                num nValue[3]
            mdesc mMdesc
            num nActionIndex = 42
            num nDelay
            num nMoveType = 1
            num nPercentage
            num nSigValue = 1
        pointRx pPointRx[2] = {x=93.576632, y=-409.183941, z=700.107773, rx=0.434495, ry=-1.660891, rz=-0.491266, shoulder=lefty, elbow=enegative, wrist=wpositive}
        string sID
      [45]
        bool bMarked
        jointRx jJointRx = {j1=-101.229016, j2=121.246473, j3=-113.173387, j4=191.93634, j5=7.483782, j6=-91.0959406}
        pointRx pInter
        paraItem pParaItem
          [0]
            bool bSafePoint
            ifItem iIfItem
              [0]
                bool bANDOR[2]
                num nSigIndex[3]
                num nSigType[3]
                num nValue[3]
            mdesc mMdesc
            num nActionIndex = 42
            num nDelay
            num nMoveType = 1
            num nPercentage
            num nSigValue = 1
        pointRx pPointRx[2] = {x=-57.556145, y=-477.506256, z=700.107677, rx=0.434341, ry=-1.659983, rz=-0.491216, shoulder=lefty, elbow=enegative, wrist=wpositive}
        string sID
      [46]
        bool bMarked
        jointRx jJointRx = {j1=-100.83359, j2=118.28296, j3=-99.234912, j4=184.924538, j5=18.376568, j6=-84.328027}
        pointRx pInter
        paraItem pParaItem
          [0]
            bool bSafePoint
            ifItem iIfItem
              [0]
                bool bANDOR[2]
                num nSigIndex[3]
                num nSigType[3]
                num nValue[3]
            mdesc mMdesc
            num nActionIndex = 42
            num nDelay
            num nMoveType = 1
            num nPercentage
            num nSigValue = 1
        pointRx pPointRx[2] = {x=-71.199798, y=-566.082474, z=700.128795, rx=0.430138, ry=-1.661253, rz=-0.490771, shoulder=lefty, elbow=enegative, wrist=wpositive}
        string sID
      [47]
        bool bMarked
        jointRx jJointRx = {j1=-96.744625, j2=116.717504, j3=-93.79165, j4=184.203052, j5=22.358435, j6=-87.631438}
        pointRx pInter
        paraItem pParaItem
          [0]
            bool bSafePoint
            ifItem iIfItem
              [0]
                bool bANDOR[2]
                num nSigIndex[3]
                num nSigType[3]
                num nValue[3]
            mdesc mMdesc
            num nActionIndex = 42
            num nDelay
            num nMoveType = 1
            num nPercentage
            num nSigValue = 1
        pointRx pPointRx[2] = {x=-34.726735, y=-600.68007, z=700.128795, rx=0.429673, ry=-1.659562, rz=-0.490424, shoulder=lefty, elbow=enegative, wrist=wpositive}
        string sID
      [48]
        bool bMarked
        jointRx jJointRx = {j1=-95.531794, j2=118.469763, j3=-99.931703, j4=185.21224, j5=18.0199205, j6=-89.914501}
        pointRx pInter
        paraItem pParaItem
          [0]
            bool bSafePoint
            ifItem iIfItem
              [0]
                bool bANDOR[2]
                num nSigIndex[3]
                num nSigType[3]
                num nValue[3]
            mdesc mMdesc
            num nActionIndex = 42
            num nDelay
            num nMoveType = 1
            num nPercentage
            num nSigValue = 1
        pointRx pPointRx[2] = {x=-18.573295, y=-564.69379, z=700.128759, rx=0.42985, ry=-1.65955, rz=-0.49045, shoulder=lefty, elbow=enegative, wrist=wpositive}
        string sID
      [49]
        bool bMarked
        jointRx jJointRx = {j1=-92.248565, j2=118.548585, j3=-100.229526, j4=185.345375, j5=17.897666, j6=-93.328956}
        pointRx pInter
        paraItem pParaItem
          [0]
            bool bSafePoint
            ifItem iIfItem
              [0]
                bool bANDOR[2]
                num nSigIndex[3]
                num nSigType[3]
                num nValue[3]
            mdesc mMdesc
            num nActionIndex = 42
            num nDelay
            num nMoveType = 1
            num nPercentage
            num nSigValue = 1
        pointRx pPointRx[2] = {x=13.638528, y=-562.185834, z=700.128755, rx=0.429526, ry=-1.658701, rz=-0.490292, shoulder=lefty, elbow=enegative, wrist=wpositive}
        string sID
      [50]
        bool bMarked
        jointRx jJointRx = {j1=-92.0110168, j2=115.175363, j3=-88.916981, j4=183.775747, j5=25.818301, j6=-91.878431}
        pointRx pInter
        paraItem pParaItem
          [0]
            bool bSafePoint
            ifItem iIfItem
              [0]
                bool bANDOR[2]
                num nSigIndex[3]
                num nSigType[3]
                num nValue[3]
            mdesc mMdesc
            num nActionIndex = 42
            num nDelay
            num nMoveType = 1
            num nPercentage
            num nSigValue = 1
        pointRx pPointRx[2] = {x=13.638517, y=-627.787273, z=700.128718, rx=0.430872, ry=-1.659586, rz=-0.490435, shoulder=lefty, elbow=enegative, wrist=wpositive}
        string sID
      [51]
        bool bMarked
        jointRx jJointRx = {j1=-97.374112, j2=108.454018, j3=-70.449442, j4=182.620747, j5=37.393534, j6=-85.196557}
        pointRx pInter
        paraItem pParaItem
          [0]
            bool bSafePoint
            ifItem iIfItem
              [0]
                bool bANDOR[2]
                num nSigIndex[3]
                num nSigType[3]
                num nValue[3]
            mdesc mMdesc
            num nActionIndex = 42
            num nDelay
            num nMoveType = 1
            num nPercentage
            num nSigValue = 1
        pointRx pPointRx[2] = {x=-56.645666, y=-719.0880848, z=700.128704, rx=0.430401, ry=-1.660167, rz=-0.490645, shoulder=lefty, elbow=enegative, wrist=wpositive}
        string sID
      [52]
        bool bMarked
        jointRx jJointRx = {j1=-97.840683, j2=111.886769, j3=-79.472132, j4=183.0096897, j5=31.798373, j6=-85.205581}
        pointRx pInter
        paraItem pParaItem
          [0]
            bool bSafePoint
            ifItem iIfItem
              [0]
                bool bANDOR[2]
                num nSigIndex[3]
                num nSigType[3]
                num nValue[3]
            mdesc mMdesc
            num nActionIndex = 42
            num nDelay
            num nMoveType = 1
            num nPercentage
            num nSigValue = 1
        pointRx pPointRx[2] = {x=-56.645667, y=-676.466244, z=700.128712, rx=0.429254, ry=-1.659449, rz=-0.490453, shoulder=lefty, elbow=enegative, wrist=wpositive}
        string sID
      [53]
        bool bMarked
        jointRx jJointRx = {j1=-99.139712, j2=112.699971, j3=-81.717312, j4=183.11065, j5=30.332067, j6=-84.0331021}
        pointRx pInter
        paraItem pParaItem
          [0]
            bool bSafePoint
            ifItem iIfItem
              [0]
                bool bANDOR[2]
                num nSigIndex[3]
                num nSigType[3]
                num nValue[3]
            mdesc mMdesc
            num nActionIndex = 42
            num nDelay
            num nMoveType = 1
            num nPercentage
            num nSigValue = 1
        pointRx pPointRx[2] = {x=-70.0879135, y=-664.155218, z=700.128714, rx=0.429183, ry=-1.659583, rz=-0.490504, shoulder=lefty, elbow=enegative, wrist=wpositive}
        string sID
      [54]
        bool bMarked
        jointRx jJointRx = {j1=-105.267989, j2=114.670594, j3=-87.395728, j4=183.340854, j5=26.462946, j6=-78.209203}
        pointRx pInter
        paraItem pParaItem
          [0]
            bool bSafePoint
            ifItem iIfItem
              [0]
                bool bANDOR[2]
                num nSigIndex[3]
                num nSigType[3]
                num nValue[3]
            mdesc mMdesc
            num nActionIndex = 42
            num nDelay
            num nMoveType = 1
            num nPercentage
            num nSigValue = 1
        pointRx pPointRx[2] = {x=-132.400518, y=-625.604431, z=700.128755, rx=0.42881, ry=-1.659576, rz=-0.490548, shoulder=lefty, elbow=enegative, wrist=wpositive}
        string sID
      [55]
        bool bMarked
        jointRx jJointRx = {j1=-104.169194, j2=109.68382, j3=-73.608878, j4=182.604541, j5=35.278725, j6=-78.44342}
        pointRx pInter
        paraItem pParaItem
          [0]
            bool bSafePoint
            ifItem iIfItem
              [0]
                bool bANDOR[2]
                num nSigIndex[3]
                num nSigType[3]
                num nValue[3]
            mdesc mMdesc
            num nActionIndex = 42
            num nDelay
            num nMoveType = 1
            num nPercentage
            num nSigValue = 1
        pointRx pPointRx[2] = {x=-137.458378, y=-695.112294, z=700.128753, rx=0.430847, ry=-1.65989, rz=-0.490478, shoulder=lefty, elbow=enegative, wrist=wpositive}
        string sID
      [56]
        bool bMarked
        jointRx jJointRx = {j1=-108.836483, j2=105.997726, j3=-64.330372, j4=182.193953, j5=40.744432, j6=-73.310916}
        pointRx pInter
        paraItem pParaItem
          [0]
            bool bSafePoint
            ifItem iIfItem
              [0]
                bool bANDOR[2]
                num nSigIndex[3]
                num nSigType[3]
                num nValue[3]
            mdesc mMdesc
            num nActionIndex = 42
            num nDelay
            num nMoveType = 1
            num nPercentage
            num nSigValue = 1
        pointRx pPointRx[2] = {x=-206.432129, y=-721.294628, z=700.128699, rx=0.4308, ry=-1.659754, rz=-0.490404, shoulder=lefty, elbow=enegative, wrist=wpositive}
        string sID
      [57]
        bool bMarked
        jointRx jJointRx = {j1=-117.384994, j2=111.318057, j3=-77.929976, j4=182.390665, j5=32.266362, j6=-65.120808}
        pointRx pInter
        paraItem pParaItem
          [0]
            bool bSafePoint
            ifItem iIfItem
              [0]
                bool bANDOR[2]
                num nSigIndex[3]
                num nSigType[3]
                num nValue[3]
            mdesc mMdesc
            num nActionIndex = 42
            num nDelay
            num nMoveType = 1
            num nPercentage
            num nSigValue = 1
        pointRx pPointRx[2] = {x=-282.767279, y=-630.359837, z=700.128774, rx=0.429, ry=-1.659295, rz=-0.490511, shoulder=lefty, elbow=enegative, wrist=wpositive}
        string sID
      [58]
        bool bMarked
        jointRx jJointRx = {j1=-126.0288968, j2=110.864642, j3=-76.715468, j4=182.00929387, j5=32.842378, j6=-56.143629}
        pointRx pInter
        paraItem pParaItem
          [0]
            bool bSafePoint
            ifItem iIfItem
              [0]
                bool bANDOR[2]
                num nSigIndex[3]
                num nSigType[3]
                num nValue[3]
            mdesc mMdesc
            num nActionIndex = 42
            num nDelay
            num nMoveType = 1
            num nPercentage
            num nSigValue = 1
        pointRx pPointRx[2] = {x=-377.367552, y=-587.693598, z=700.128774, rx=0.428889, ry=-1.659196, rz=-0.49055, shoulder=lefty, elbow=enegative, wrist=wpositive}
        string sID
      [59]
        bool bMarked
        jointRx jJointRx = {j1=-132.158352, j2=110.822497, j3=-76.606813, j4=181.740658, j5=32.799901, j6=-49.794511}
        pointRx pInter
        paraItem pParaItem
          [0]
            bool bSafePoint
            ifItem iIfItem
              [0]
                bool bANDOR[2]
                num nSigIndex[3]
                num nSigType[3]
                num nValue[3]
            mdesc mMdesc
            num nActionIndex = 42
            num nDelay
            num nMoveType = 1
            num nPercentage
            num nSigValue = 1
        pointRx pPointRx[2] = {x=-437.975867, y=-545.96373, z=700.144476, rx=0.425586, ry=-1.657208, rz=-0.495183, shoulder=lefty, elbow=enegative, wrist=wpositive}
        string sID
      [60]
        bool bMarked
        jointRx jJointRx = {j1=-130.472656, j2=91.957177, j3=-58.182906, j4=181.836817, j5=32.386471, j6=-51.5677}
        pointRx pInter
        paraItem pParaItem
          [0]
            bool bSafePoint
            ifItem iIfItem
              [0]
                bool bANDOR[2]
                num nSigIndex[3]
                num nSigType[3]
                num nValue[3]
            mdesc mMdesc
            num nActionIndex = 42
            num nDelay
            num nMoveType = 1
            num nPercentage
            num nSigValue = 1
        pointRx pPointRx[2] = {x=-437.940696, y=-577.0648472, z=838.536537, rx=0.42728, ry=-1.657753, rz=-0.494943, shoulder=lefty, elbow=enegative, wrist=wpositive}
        string sID
      [61]
        bool bMarked
        jointRx jJointRx = {j1=-136.0523069, j2=93.884763, j3=-71.42598, j4=182.356, j5=20.985823, j6=-46.637919}
        pointRx pInter
        paraItem pParaItem
          [0]
            bool bSafePoint
            ifItem iIfItem
              [0]
                bool bANDOR[2]
                num nSigIndex[3]
                num nSigType[3]
                num nValue[3]
            mdesc mMdesc
            num nActionIndex = 42
            num nDelay
            num nMoveType = 1
            num nPercentage
            num nSigValue = 1
        pointRx pPointRx[2] = {x=-437.940746, y=-481.365195, z=863.748923, rx=0.426109, ry=-1.657561, rz=-0.495141, shoulder=lefty, elbow=enegative, wrist=wpositive}
        string sID
      [62]
        bool bMarked
        jointRx jJointRx = {j1=-136.052274, j2=115.42016, j3=-86.959194, j4=181.859406, j5=26.985128, j6=-46.0951129}
        pointRx pInter
        paraItem pParaItem
          [0]
            bool bSafePoint
            ifItem iIfItem
              [0]
                bool bANDOR[2]
                num nSigIndex[3]
                num nSigType[3]
                num nValue[3]
            mdesc mMdesc
            num nActionIndex = 42
            num nDelay
            num nMoveType = 1
            num nPercentage
            num nSigValue = 1
        pointRx pPointRx[2] = {x=-437.940805, y=-481.365263, z=690.980039, rx=0.425304, ry=-1.656785, rz=-0.495111, shoulder=lefty, elbow=enegative, wrist=wpositive}
        string sID
      [63]
        bool bMarked
        jointRx jJointRx = {j1=-87.550712, j2=145.128314, j3=-83.0892372, j4=182.118111, j5=63.690986, j6=-64.966608}
        pointRx pInter
        paraItem pParaItem
          [0]
            bool bSafePoint
            ifItem iIfItem
              [0]
                bool bANDOR[2]
                num nSigIndex[3]
                num nSigType[3]
                num nValue[3]
            mdesc mMdesc
            num nActionIndex = 42
            num nDelay
            num nMoveType = 1
            num nPercentage
            num nSigValue = 1
        pointRx pPointRx[2] = {x=61.357264, y=-652.082, z=350.106484, rx=-1.553715, ry=-1.966811, rz=28.422241, shoulder=lefty, elbow=enegative, wrist=wpositive}
        string sID
    string sID
  [Position6_point_wash]
    num nFrameIndex
    num nMoveID
    num nToolIndex
    pointItem pPointItem[65]
      [0]
        bool bMarked
        jointRx jJointRx
        pointRx pInter
        paraItem pParaItem
          [0]
            bool bSafePoint
            ifItem iIfItem
              [0]
                bool bANDOR[2]
                num nSigIndex[3]
                num nSigType[3]
                num nValue[3]
            mdesc mMdesc
            num nActionIndex = 41
            num nDelay
            num nMoveType = 4
            num nPercentage
            num nSigValue = 1
        pointRx pPointRx[2]
        string sID
      [1]
        bool bMarked
        jointRx jJointRx
        pointRx pInter
        paraItem pParaItem
          [0]
            bool bSafePoint
            ifItem iIfItem
              [0]
                bool bANDOR[2]
                num nSigIndex[3]
                num nSigType[3]
                num nValue[3]
            mdesc mMdesc
            num nActionIndex = 42
            num nDelay
            num nMoveType = 4
            num nPercentage
            num nSigValue = 1
        pointRx pPointRx[2]
        string sID
      [2]
        bool bMarked
        jointRx jJointRx = {j1=-87.550712, j2=145.128314, j3=-83.0892365, j4=182.11811, j5=63.690987, j6=-64.966608}
        pointRx pInter
        paraItem pParaItem
          [0]
            bool bSafePoint
            ifItem iIfItem
              [0]
                bool bANDOR[2]
                num nSigIndex[3]
                num nSigType[3]
                num nValue[3]
            mdesc mMdesc
            num nActionIndex = 42
            num nDelay
            num nMoveType = 1
            num nPercentage
            num nSigValue = 1
        pointRx pPointRx[2] = {x=61.357264, y=-652.082, z=350.106484, rx=-1.553715, ry=-1.966811, rz=28.422241, shoulder=lefty, elbow=enegative, wrist=wpositive}
        string sID
      [3]
        bool bMarked
        jointRx jJointRx = {j1=-58.982134, j2=104.832128, j3=-61.565333, j4=183.343645, j5=42.668286, j6=-33.606181}
        pointRx pInter
        paraItem pParaItem
          [0]
            bool bSafePoint
            ifItem iIfItem
              [0]
                bool bANDOR[2]
                num nSigIndex[3]
                num nSigType[3]
                num nValue[3]
            mdesc mMdesc
            num nActionIndex = 42
            num nDelay
            num nMoveType = 1
            num nPercentage
            num nSigValue = 1
        pointRx pPointRx[2] = {x=416.397495, y=-633.838238, z=700.254781, rx=1.722211, ry=-1.608013, rz=89.88289, shoulder=lefty, elbow=enegative, wrist=wpositive}
        string sID
      [4]
        bool bMarked
        jointRx jJointRx = {j1=-62.332645, j2=107.50753, j3=-68.132801, j4=183.562396, j5=38.651057, j6=-30.577163}
        pointRx pInter
        paraItem pParaItem
          [0]
            bool bSafePoint
            ifItem iIfItem
              [0]
                bool bANDOR[2]
                num nSigIndex[3]
                num nSigType[3]
                num nValue[3]
            mdesc mMdesc
            num nActionIndex = 42
            num nDelay
            num nMoveType = 1
            num nPercentage
            num nSigValue = 1
        pointRx pPointRx[2] = {x=366.85786, y=-633.838275, z=700.254798, rx=1.721666, ry=-1.608681, rz=89.88277, shoulder=lefty, elbow=enegative, wrist=wpositive}
        string sID
      [5]
        bool bMarked
        jointRx jJointRx = {j1=-67.0327916, j2=110.2281, j3=-75.107293, j4=183.830258, j5=34.223084, j6=-26.259259}
        pointRx pInter
        paraItem pParaItem
          [0]
            bool bSafePoint
            ifItem iIfItem
              [0]
                bool bANDOR[2]
                num nSigIndex[3]
                num nSigType[3]
                num nValue[3]
            mdesc mMdesc
            num nActionIndex = 42
            num nDelay
            num nMoveType = 1
            num nPercentage
            num nSigValue = 1
        pointRx pPointRx[2] = {x=302.522929, y=-633.83826, z=700.254794, rx=1.721622, ry=-1.608914, rz=89.882692, shoulder=lefty, elbow=enegative, wrist=wpositive}
        string sID
      [6]
        bool bMarked
        jointRx jJointRx = {j1=-71.633736, j2=112.694899, j3=-81.788319, j4=184.160101, j5=29.845031, j6=-22.0972061}
        pointRx pInter
        paraItem pParaItem
          [0]
            bool bSafePoint
            ifItem iIfItem
              [0]
                bool bANDOR[2]
                num nSigIndex[3]
                num nSigType[3]
                num nValue[3]
            mdesc mMdesc
            num nActionIndex = 42
            num nDelay
            num nMoveType = 1
            num nPercentage
            num nSigValue = 1
        pointRx pPointRx[2] = {x=241.500206, y=-626.00943449, z=700.254792, rx=1.721289, ry=-1.608551, rz=89.882813, shoulder=lefty, elbow=enegative, wrist=wpositive}
        string sID
      [7]
        bool bMarked
        jointRx jJointRx = {j1=-65.27374, j2=114.413405, j3=-86.726434, j4=184.827216, j5=26.876761, j6=-29.158228}
        pointRx pInter
        paraItem pParaItem
          [0]
            bool bSafePoint
            ifItem iIfItem
              [0]
                bool bANDOR[2]
                num nSigIndex[3]
                num nSigType[3]
                num nValue[3]
            mdesc mMdesc
            num nActionIndex = 42
            num nDelay
            num nMoveType = 1
            num nPercentage
            num nSigValue = 1
        pointRx pPointRx[2] = {x=296.78184, y=-570.410131, z=700.254763, rx=1.722456, ry=-1.607129, rz=89.88308, shoulder=lefty, elbow=enegative, wrist=wpositive}
        string sID
      [8]
        bool bMarked
        jointRx jJointRx = {j1=-60.709616, j2=114.554511, j3=-87.145192, j4=184.986355, j5=26.782513, j6=-33.871303}
        pointRx pInter
        paraItem pParaItem
          [0]
            bool bSafePoint
            ifItem iIfItem
              [0]
                bool bANDOR[2]
                num nSigIndex[3]
                num nSigType[3]
                num nValue[3]
            mdesc mMdesc
            num nActionIndex = 42
            num nDelay
            num nMoveType = 1
            num nPercentage
            num nSigValue = 1
        pointRx pPointRx[2] = {x=338.875527, y=-541.934118, z=700.254791, rx=1.721113, ry=-1.608268, rz=89.882966, shoulder=lefty, elbow=enegative, wrist=wpositive}
        string sID
      [9]
        bool bMarked
        jointRx jJointRx = {j1=-66.643474, j2=118.657481, j3=-100.787497, j4=187.380827, j5=17.0599953, j6=-30.539636}
        pointRx pInter
        paraItem pParaItem
          [0]
            bool bSafePoint
            ifItem iIfItem
              [0]
                bool bANDOR[2]
                num nSigIndex[3]
                num nSigType[3]
                num nValue[3]
            mdesc mMdesc
            num nActionIndex = 42
            num nDelay
            num nMoveType = 1
            num nPercentage
            num nSigValue = 1
        pointRx pPointRx[2] = {x=251.241513, y=-503.208169, z=700.254788, rx=1.722301, ry=-1.608953, rz=89.882703, shoulder=lefty, elbow=enegative, wrist=wpositive}
        string sID
      [10]
        bool bMarked
        jointRx jJointRx = {j1=-65.0394334, j2=119.495527, j3=-104.191107, j4=188.704216, j5=14.582841, j6=-33.512784}
        pointRx pInter
        paraItem pParaItem
          [0]
            bool bSafePoint
            ifItem iIfItem
              [0]
                bool bANDOR[2]
                num nSigIndex[3]
                num nSigType[3]
                num nValue[3]
            mdesc mMdesc
            num nActionIndex = 42
            num nDelay
            num nMoveType = 1
            num nPercentage
            num nSigValue = 1
        pointRx pPointRx[2] = {x=255.846551, y=-476.313024, z=700.254767, rx=1.721654, ry=-1.607307, rz=89.883015, shoulder=lefty, elbow=enegative, wrist=wpositive}
        string sID
      [11]
        bool bMarked
        jointRx jJointRx = {j1=-71.0596735, j2=121.00750191, j3=-111.877772, j4=194.578806, j5=8.286602, j6=-33.494479}
        pointRx pInter
        paraItem pParaItem
          [0]
            bool bSafePoint
            ifItem iIfItem
              [0]
                bool bANDOR[2]
                num nSigIndex[3]
                num nSigType[3]
                num nValue[3]
            mdesc mMdesc
            num nActionIndex = 42
            num nDelay
            num nMoveType = 1
            num nPercentage
            num nSigValue = 1
        pointRx pPointRx[2] = {x=189.620191, y=-454.405925, z=700.254767, rx=1.721353, ry=-1.607377, rz=89.882905, shoulder=lefty, elbow=enegative, wrist=wpositive}
        string sID
      [12]
        bool bMarked
        jointRx jJointRx = {j1=-74.809464, j2=121.0382904, j3=-112.0769955, j4=194.59856, j5=7.974501, j6=-29.773551}
        pointRx pInter
        paraItem pParaItem
          [0]
            bool bSafePoint
            ifItem iIfItem
              [0]
                bool bANDOR[2]
                num nSigIndex[3]
                num nSigType[3]
                num nValue[3]
            mdesc mMdesc
            num nActionIndex = 42
            num nDelay
            num nMoveType = 1
            num nPercentage
            num nSigValue = 1
        pointRx pPointRx[2] = {x=160.082647, y=-465.491863, z=700.254784, rx=1.722803, ry=-1.608682, rz=89.882806, shoulder=lefty, elbow=enegative, wrist=wpositive}
        string sID
      [13]
        bool bMarked
        jointRx jJointRx = {j1=-76.815291, j2=120.680634, j3=-109.926019, j4=191.777648, j5=9.643692, j6=-24.919524}
        pointRx pInter
        paraItem pParaItem
          [0]
            bool bSafePoint
            ifItem iIfItem
              [0]
                bool bANDOR[2]
                num nSigIndex[3]
                num nSigType[3]
                num nValue[3]
            mdesc mMdesc
            num nActionIndex = 42
            num nDelay
            num nMoveType = 1
            num nPercentage
            num nSigValue = 1
        pointRx pPointRx[2] = {x=147.50556, y=-485.393693, z=700.254789, rx=1.722658, ry=-1.609045, rz=89.882735, shoulder=lefty, elbow=enegative, wrist=wpositive}
        string sID
      [14]
        bool bMarked
        jointRx jJointRx = {j1=-80.979539, j2=121.627826, j3=-116.887787, j4=209.4559, j5=3.779386, j6=-38.540773}
        pointRx pInter
        paraItem pParaItem
          [0]
            bool bSafePoint
            ifItem iIfItem
              [0]
                bool bANDOR[2]
                num nSigIndex[3]
                num nSigType[3]
                num nValue[3]
            mdesc mMdesc
            num nActionIndex = 42
            num nDelay
            num nMoveType = 1
            num nPercentage
            num nSigValue = 1
        pointRx pPointRx[2] = {x=105.438294, y=-448.641412, z=700.254346, rx=1.721348, ry=-1.60753, rz=89.882882, shoulder=lefty, elbow=enegative, wrist=wpositive}
        string sID
      [15]
        bool bMarked
        jointRx jJointRx = {j1=-97.0735787, j2=120.583034, j3=-109.386983, j4=169.0121648, j5=9.967554, j6=107.0502076}
        pointRx pInter
        paraItem pParaItem
          [0]
            bool bSafePoint
            ifItem iIfItem
              [0]
                bool bANDOR[2]
                num nSigIndex[3]
                num nSigType[3]
                num nValue[3]
            mdesc mMdesc
            num nActionIndex = 42
            num nDelay
            num nMoveType = 1
            num nPercentage
            num nSigValue = 1
        pointRx pPointRx[2] = {x=3.102788, y=-514.97816, z=700.254373, rx=1.629756, ry=1.702884, rz=179.149702, shoulder=lefty, elbow=enegative, wrist=wpositive}
        string sID
      [16]
        bool bMarked
        jointRx jJointRx = {j1=-98.785966, j2=121.589944, j3=-116.474742, j4=152.822693, j5=4.230949, j6=125.0509123}
        pointRx pInter
        paraItem pParaItem
          [0]
            bool bSafePoint
            ifItem iIfItem
              [0]
                bool bANDOR[2]
                num nSigIndex[3]
                num nSigType[3]
                num nValue[3]
            mdesc mMdesc
            num nActionIndex = 42
            num nDelay
            num nMoveType = 1
            num nPercentage
            num nSigValue = 1
        pointRx pPointRx[2] = {x=-4.455751, y=-466.481228, z=700.254288, rx=1.629056, ry=1.702249, rz=179.149669, shoulder=lefty, elbow=enegative, wrist=wpositive}
        string sID
      [17]
        bool bMarked
        jointRx jJointRx = {j1=-102.289362, j2=121.662055, j3=-117.287244, j4=147.396601, j5=3.732456, j6=133.989908}
        pointRx pInter
        paraItem pParaItem
          [0]
            bool bSafePoint
            ifItem iIfItem
              [0]
                bool bANDOR[2]
                num nSigIndex[3]
                num nSigType[3]
                num nValue[3]
            mdesc mMdesc
            num nActionIndex = 42
            num nDelay
            num nMoveType = 1
            num nPercentage
            num nSigValue = 1
        pointRx pPointRx[2] = {x=-30.830703, y=-458.833227, z=700.253116, rx=1.628925, ry=1.702444, rz=179.149706, shoulder=lefty, elbow=enegative, wrist=wpositive}
        string sID
      [18]
        bool bMarked
        jointRx jJointRx = {j1=-97.596795, j2=121.636094, j3=-116.996972, j4=154.0724475, j5=5.372504, j6=163.484863}
        pointRx pInter
        paraItem pParaItem
          [0]
            bool bSafePoint
            ifItem iIfItem
              [0]
                bool bANDOR[2]
                num nSigIndex[3]
                num nSigType[3]
                num nValue[3]
            mdesc mMdesc
            num nActionIndex = 42
            num nDelay
            num nMoveType = 1
            num nPercentage
            num nSigValue = 1
        pointRx pPointRx[2] = {x=11.0855283, y=-449.928798, z=700.263578, rx=0.116735, ry=2.351476, rz=-139.946822, shoulder=lefty, elbow=enegative, wrist=wpositive}
        string sID
      [19]
        bool bMarked
        jointRx jJointRx = {j1=-93.435678, j2=120.973902, j3=-111.67187, j4=165.758899, j5=9.616057, j6=147.540776}
        pointRx pInter
        paraItem pParaItem
          [0]
            bool bSafePoint
            ifItem iIfItem
              [0]
                bool bANDOR[2]
                num nSigIndex[3]
                num nSigType[3]
                num nValue[3]
            mdesc mMdesc
            num nActionIndex = 42
            num nDelay
            num nMoveType = 1
            num nPercentage
            num nSigValue = 1
        pointRx pPointRx[2] = {x=41.481677, y=-486.244692, z=700.26363, rx=0.117474, ry=2.35234, rz=-139.946783, shoulder=lefty, elbow=enegative, wrist=wpositive}
        string sID
      [20]
        bool bMarked
        jointRx jJointRx = {j1=-87.514361, j2=121.638618, j3=-117.0243701, j4=151.901605, j5=4.980778, j6=155.573887}
        pointRx pInter
        paraItem pParaItem
          [0]
            bool bSafePoint
            ifItem iIfItem
              [0]
                bool bANDOR[2]
                num nSigIndex[3]
                num nSigType[3]
                num nValue[3]
            mdesc mMdesc
            num nActionIndex = 42
            num nDelay
            num nMoveType = 1
            num nPercentage
            num nSigValue = 1
        pointRx pPointRx[2] = {x=89.805675, y=-444.448305, z=700.262762, rx=0.116151, ry=2.350833, rz=-139.946826, shoulder=lefty, elbow=enegative, wrist=wpositive}
        string sID
      [21]
        bool bMarked
        jointRx jJointRx = {j1=-85.538373, j2=121.159338, j3=-112.89672, j4=163.596021, j5=8.296682, j6=141.829296}
        pointRx pInter
        paraItem pParaItem
          [0]
            bool bSafePoint
            ifItem iIfItem
              [0]
                bool bANDOR[2]
                num nSigIndex[3]
                num nSigType[3]
                num nValue[3]
            mdesc mMdesc
            num nActionIndex = 42
            num nDelay
            num nMoveType = 1
            num nPercentage
            num nSigValue = 1
        pointRx pPointRx[2] = {x=107.297774, y=-470.450865, z=700.262819, rx=0.116544, ry=2.351714, rz=-139.94676, shoulder=lefty, elbow=enegative, wrist=wpositive}
        string sID
      [22]
        bool bMarked
        jointRx jJointRx = {j1=-80.389938, j2=121.305327, j3=-113.961147, j4=161.375696, j5=7.211507, j6=138.92232}
        pointRx pInter
        paraItem pParaItem
          [0]
            bool bSafePoint
            ifItem iIfItem
              [0]
                bool bANDOR[2]
                num nSigIndex[3]
                num nSigType[3]
                num nValue[3]
            mdesc mMdesc
            num nActionIndex = 42
            num nDelay
            num nMoveType = 1
            num nPercentage
            num nSigValue = 1
        pointRx pPointRx[2] = {x=147.836969, y=-453.554332, z=700.262491, rx=0.115759, ry=2.349936, rz=-139.946858, shoulder=lefty, elbow=enegative, wrist=wpositive}
        string sID
      [23]
        bool bMarked
        jointRx jJointRx = {j1=-74.160542, j2=121.48868, j3=-115.480429, j4=163.296331, j5=4.15176, j6=89.975533}
        pointRx pInter
        paraItem pParaItem
          [0]
            bool bSafePoint
            ifItem iIfItem
              [0]
                bool bANDOR[2]
                num nSigIndex[3]
                num nSigType[3]
                num nValue[3]
            mdesc mMdesc
            num nActionIndex = 42
            num nDelay
            num nMoveType = 1
            num nPercentage
            num nSigValue = 1
        pointRx pPointRx[2] = {x=187.654652, y=-440.110471, z=700.252779, rx=1.628669, ry=1.701382, rz=179.149675, shoulder=lefty, elbow=enegative, wrist=wpositive}
        string sID
      [24]
        bool bMarked
        jointRx jJointRx = {j1=-69.509661, j2=119.265921, j3=-103.220112, j4=175.749132, j5=13.961301, j6=72.790426}
        pointRx pInter
        paraItem pParaItem
          [0]
            bool bSafePoint
            ifItem iIfItem
              [0]
                bool bANDOR[2]
                num nSigIndex[3]
                num nSigType[3]
                num nValue[3]
            mdesc mMdesc
            num nActionIndex = 42
            num nDelay
            num nMoveType = 1
            num nPercentage
            num nSigValue = 1
        pointRx pPointRx[2] = {x=250.0960558, y=-500.875002, z=700.252775, rx=1.628687, ry=1.702386, rz=179.149806, shoulder=lefty, elbow=enegative, wrist=wpositive}
        string sID
      [25]
        bool bMarked
        jointRx jJointRx = {j1=-65.451313, j2=120.0346612, j3=-106.615882, j4=175.540521, j5=11.264344, j6=68.982362}
        pointRx pInter
        paraItem pParaItem
          [0]
            bool bSafePoint
            ifItem iIfItem
              [0]
                bool bANDOR[2]
                num nSigIndex[3]
                num nSigType[3]
                num nValue[3]
            mdesc mMdesc
            num nActionIndex = 42
            num nDelay
            num nMoveType = 1
            num nPercentage
            num nSigValue = 1
        pointRx pPointRx[2] = {x=274.930404, y=-463.298611, z=700.25277, rx=1.6286, ry=1.700384, rz=179.149585, shoulder=lefty, elbow=enegative, wrist=wpositive}
        string sID
      [26]
        bool bMarked
        jointRx jJointRx = {j1=-63.0913911, j2=120.463088, j3=-108.745441, j4=175.274971, j5=9.527094, j6=66.910352}
        pointRx pInter
        paraItem pParaItem
          [0]
            bool bSafePoint
            ifItem iIfItem
              [0]
